(* IEC 61131-3 sources: NachHouse_TST/API/api_V12 (part 2) *)

(* ---- _07_RxBuf.ST ---- *)
// Limity jedného prijímacieho bloku a celého súboru ; Limits for one receive block and the complete file.
VAR_GLOBAL CONSTANT
  RB_BYTES {HIDDEN}    : UINT := 256;     // Maximálny počet dátových bajtov v jednom bloku ; Maximum data bytes in one block.
  RB_FILE_MAX {HIDDEN} : UDINT := 65535;  // Maximálna veľkosť súboru, ktorý možno zložiť ; Maximum size of a file that can be assembled.
END_VAR

VAR_GLOBAL
  RbSeen     : UDINT := 0;            // Posledná požiadavka bloku už prijatá PLC ; Most recent block request already consumed by the PLC.
  RbActive   : BOOL := FALSE;         // TRUE počas skladania viacerých blokov jedného súboru ; TRUE while assembling a file from multiple blocks.
  RbTotalW   : UDINT := 0;            // Očakávaná celková dĺžka aktuálneho súboru ; Expected total length of the current file.
  RbCrcW     : DWORD := 0;            // Očakávaný CRC32 súčet aktuálneho súboru ; Expected CRC32 checksum for the current file.
  RbCrcState : DWORD := 16#FFFFFFFF;  // Medzistav výpočtu CRC32 medzi prijatými blokmi ; Running CRC32 state across received blocks.
END_VAR

// Jeden krok štandardného CRC32 pre jeden bajt ; polynóm je 0xEDB88320. ; One standard CRC32 step for a byte ; the polynomial is 0xEDB88320.
// Pridá jeden bajt do priebežného výpočtu CRC32 ; Add one byte to the running CRC32 calculation.
FUNCTION RbCrcByte : DWORD
  VAR_INPUT
    State : DWORD;  // Doterajší priebežný stav CRC ; Previous running CRC state.
    B     : BYTE;   // Bajt, ktorý sa pridáva do CRC ; Byte to add to the CRC.
  END_VAR
  VAR
    C : DWORD;  // Pracovný 32-bitový stav CRC ; Working 32-bit CRC value.
    I : USINT;  // Počet ôsmich bitových krokov jedného bajtu ; Counter for the eight bit steps of one byte.
  END_VAR
  C := State XOR BYTE_TO_DWORD(B);
  FOR I := 1 TO 8 DO
    IF (C AND 16#00000001) <> 0 THEN
      C := SHR(C, 1) XOR 16#EDB88320;
    ELSE
      C := SHR(C, 1);
    END_IF;
  END_FOR;
  RbCrcByte := C;
END_FUNCTION

// Každé nové RbRq spracuje jeden blok ; RbAck potvrdí spracovanie a RbErr výsledok. ; Each new RbRq processes one block ; RbAck acknowledges it and RbErr reports the result.
// RbReady sa nastaví až po kontrole veľkosti a CRC celého súboru. ; RbReady is set only after validating the full file size and CRC.
// Pri novej RbRq zapíše jeden blok do rx.json, priebežne počíta CRC a potvrdí výsledok ; On a new RbRq, write one block to rx.json, update CRC, and acknowledge the result.
FUNCTION RbCycle : BOOL
  VAR
    Hnd      : HANDLE;       // Otvorený súborový handle pre zápis bloku ; File handle used to write the block.
    Mode     : TF_MODE;      // Režim otvorenia: nový súbor alebo pripojenie ďalšieho bloku ; Open mode: create a file or append the next block.
    N        : UDINT;        // Počet bajtov, ktoré FileWrite skutočne zapísal ; Number of bytes actually written by FileWrite.
    I        : UINT;         // Index bajtu pri aktualizácii CRC ; Byte index while updating the CRC.
    PB       : PTR_TO BYTE;  // Ukazovateľ na postupné čítanie bajtov z rxBuf ; Pointer used to read bytes sequentially from rxBuf.
    Closed   : BOOL;         // Výsledok uzatvorenia súboru po zápise ; Result of closing the file after writing.
    FinalCrc : DWORD;        // Dokončený CRC32 súčet po spracovaní posledného bajtu ; Final CRC32 value after the last byte.
  END_VAR
  RbCycle := TRUE;
  // Bez nového čísla požiadavky sa blok nespracúva znova ; Do not process a block again without a new request number.
  IF (RbRq = 0) OR (RbRq = RbSeen) THEN RETURN; END_IF;
  RbSeen := RbRq;
  RbErr := 0;

  // Počas parsovania JSON-u sa ďalší blok odmietne, aby sa súbor nemenil pod parserom ; Reject a new block while JSON parsing is active so the file cannot change underneath the parser.
  IF RxSt <> 0 THEN RbErr := 10;
  ELSIF (RbLen = 0) OR (RbLen > RB_BYTES) THEN RbErr := 1;
  ELSIF (RbTotal = 0) OR (RbTotal > RB_FILE_MAX) THEN RbErr := 2;
  ELSIF RbOfs > RbTotal THEN RbErr := 3;
  ELSIF UINT_TO_UDINT(RbLen) > RbTotal - RbOfs THEN RbErr := 3;
  END_IF;

  // Pokračuje iba po úspešných kontrolách dĺžky a rozsahu ; Continue only after length and range validation succeeds.
  IF RbErr = 0 THEN
    IF RbOfs = 0 THEN
      RbActive := TRUE;
      RbReady := FALSE;
      RbWrote := 0;
      RbTotalW := RbTotal;
      RbCrcW := RbCrc;
      RbCrcState := 16#FFFFFFFF;
      Mode := F_WRITE;
    ELSE
      Mode := F_APPEND;
      IF NOT RbActive THEN RbErr := 4;
      ELSIF RbOfs <> RbWrote THEN RbErr := 5;
      ELSIF (RbTotal <> RbTotalW) OR (RbCrc <> RbCrcW) THEN RbErr := 6;
      END_IF;
    END_IF;
  END_IF;

  // Pokračuje iba po úspešných kontrolách dĺžky a rozsahu ; Continue only after length and range validation succeeds.
  IF RbErr = 0 THEN
    Hnd := FileOpen(fileName := RxPath, mode := Mode);  // Otvorí rx.json na prvý zápis alebo doplnenie bloku ; Open rx.json for the first write or for appending a block.
    IF Hnd = INVALID_HANDLE_VALUE THEN
      RbErr := 7;
      RbActive := FALSE;
    ELSE
      N := FileWrite(hFile := Hnd, adrBuf := PTR_TO_UDINT(ADR(rxBuf[0])),
                     size := UINT_TO_UDINT(RbLen));
      Closed := FileClose(hFile := Hnd);
      IF (N <> UINT_TO_UDINT(RbLen)) OR NOT Closed THEN
        RbErr := 8;
        RbActive := FALSE;
      ELSE
        PB := ADR(rxBuf[0]);  // Začne kontrolný súčet od prvého bajtu aktuálneho bloku ; Start checksum calculation at the first byte of this block.
        FOR I := 1 TO RbLen DO
          RbCrcState := RbCrcByte(State := RbCrcState, B := PB^);
          PB := UDINT_TO_PTR(PTR_TO_UDINT(PB) + 1);
        END_FOR;
        RbWrote := RbWrote + UINT_TO_UDINT(RbLen);
        // Po prijatí deklarovaného počtu bajtov overí CRC celého súboru ; Once the declared byte count arrives, verify the complete-file CRC.
        IF RbWrote = RbTotalW THEN
          FinalCrc := RbCrcState XOR 16#FFFFFFFF;
          IF FinalCrc = RbCrcW THEN
            RbReady := TRUE;
          ELSE
            RbErr := 9;
          END_IF;
          RbActive := FALSE;
        END_IF;
      END_IF;
    END_IF;
  END_IF;

  RbAck := RbRq;  // Potvrdí spracovanie aj prípadnú chybu tohto bloku ; Acknowledge processing, including any block error.
  RbCycle := RbErr = 0;
END_FUNCTION

(* ---- _02_DataInit.ST ---- *)
// Naplní testovacie záznamy a jednorazovo ich skopíruje do mRam. ; Populate test records and copy them into mRam once.
// Pri prvom cykle vytvorí testovacie ROOM/USER dáta a skopíruje ich do mRam ; On the first cycle, creates test ROOM/USER data and copies it into mRam.
FUNCTION InitData : BOOL
  VAR
    Rec    : INT;    // Index testovanej vety 1..10 ; Test record index, 1..10.
    Pos    : INT;    // Index prvku vnútorného poľa používateľa ; Index into a nested user array.
    Copied : UDINT;  // Počet bajtov skutočne skopírovaných funkciou MemCpyPtr ; Number of bytes actually copied by MemCpyPtr.
  END_VAR
  InitData := TRUE;
  // Inicializáciu vykoná iba pri štartovacej hodnote Ini ; Initialize only when Ini has its startup value.
  IF aSys.Ini <> 250 THEN RETURN; END_IF;

  // Naplnenie desiatich testovacích viet oboch typov ; Fill ten test records for both data types.
  FOR Rec := 1 TO 10 DO
    yRooms[Rec].mem.rec.Ok := TRUE;  // Začiatok naplnenia stavovej a konfiguračnej časti aktuálnej miestnosti ; Begin filling the current room's state and configuration.
    yRooms[Rec].mem.rec.ID := Rec;
    yRooms[Rec].mem.all.RoomID := Rec;
    yRooms[Rec].mem.all.CategoryID := 5;
    yRooms[Rec].mem.Temperature := 20.0 + INT_TO_REAL(Rec);
    yRooms[Rec].mem.Humidity := 40.0 + INT_TO_REAL(Rec);
    yRooms[Rec].mem.Presence := (Rec MOD 2) = 0;
    yRooms[Rec].mem.DayPhase := INT_TO_UINT(140 + Rec);
    yRooms[Rec].mem.CategoryMask := 16#00000005;
    yRooms[Rec].mem.AlarmLevel := INT_TO_USINT(Rec MOD 3);
    yRooms[Rec].mem.Online := TRUE;
    yRooms[Rec].mem.Twilight := (Rec MOD 2) <> 0;
    yRooms[Rec].cfg.Name := 'Test room';
    yRooms[Rec].cfg._Dint := INT_TO_DINT(-1000 - Rec);
    yRooms[Rec].cfg._Sint := INT_TO_SINT(-10 + Rec);
    yRooms[Rec].cfg._Usint := INT_TO_USINT(100 + Rec);
    yRooms[Rec].cfg._Uint := INT_TO_UINT(1000 + Rec);
    yRooms[Rec].cfg._Real := 10.5 + INT_TO_REAL(Rec);
    yRooms[Rec].cfg._LReal := 1000.5 + INT_TO_LREAL(Rec);
    yRooms[Rec].cfg._String := '';
    yRooms[Rec].cfg._StringCZSK := 'SVKBEGIN_+ľščťžýáíé_SVKEND';
    yRooms[Rec].cfg._BYTE := 16#A5; yRooms[Rec].cfg._WORD := 16#A55A;
    yRooms[Rec].cfg._TIME := T#12h34m56s789ms;
    yRooms[Rec].cfg._DATE := D#2026-10-07;
    yRooms[Rec].cfg._TIME_OF_DAY := TOD#12:34:56.789;
    yRooms[Rec].cfg._DATE_AND_TIME := DT#2026-10-07-12:34:56.789;

    yUsers[Rec].mem.rec.Ok := TRUE; yUsers[Rec].mem.rec.ID := Rec;  // Začiatok naplnenia aktuálnej testovacej vety USER ; Begin filling the current USER test record.
    yUsers[Rec].mem.all.RoomID := Rec; yUsers[Rec].mem.all.CategoryID := 1;
    yUsers[Rec].mem.Connected := (Rec MOD 2) = 0;
    yUsers[Rec].mem.LastError := '';
    yUsers[Rec].mem.LastUpdate := UDINT#2026100700 + INT_TO_UDINT(Rec);
    yUsers[Rec].cfg.Name := 'Test user'; yUsers[Rec].cfg.LoginHome := TRUE;
    yUsers[Rec].cfg.DshSet := FALSE; yUsers[Rec].cfg.OwnDSH := TRUE;
    yUsers[Rec].cfg.OwnQCK := TRUE;
    yUsers[Rec].cfg.UsrRight := INT_TO_USINT(1 + (Rec MOD 3));
    // Zónové oprávnenia sa menia podľa čísla testovacej vety ; Zone permissions vary with the test-record number.
    FOR Pos := 1 TO 16 DO yUsers[Rec].cfg.ZonList[Pos] := Pos <= (Rec + 1); END_FOR;
    yUsers[Rec].cfg.sbj := INT_TO_USINT(Rec);
    yUsers[Rec].cfg.lng := INT_TO_USINT(Rec MOD 2);
    FOR Pos := 0 TO 7 DO
      yUsers[Rec].cfg.fav[Pos] := INT_TO_USINT(Pos + Rec);
      yUsers[Rec].cfg.msg[Pos] := Pos = (Rec MOD 8);
    END_FOR;
    yUsers[Rec].cfg.keyPas := '123456'; yUsers[Rec].cfg.IPnbr := 1;
    yUsers[Rec].cfg.IP[1] := '192.168.33.10';
    yUsers[Rec].cfg.IP[2] := ''; yUsers[Rec].cfg.IP[3] := '';
    yUsers[Rec].cfg.mail := 'test@example.com';
    yUsers[Rec].cfg.TOKENAPPLE := 'apple-test-token';
    yUsers[Rec].cfg.TOKENUNI := 'uni-test-token';
    yUsers[Rec].cfg.gsm := '+421900000000';
    yUsers[Rec].cfg.skin := INT_TO_USINT(Rec MOD 2);
    FOR Pos := 0 TO 30 DO
      IF Pos = 0 THEN yUsers[Rec].cfg.Brw[Pos] := 0;
      ELSE yUsers[Rec].cfg.Brw[Pos] := 1;
      END_IF;
    END_FOR;
  END_FOR;

  aCfg[1].iRam := 0;  // ROOM zaberá prvú oblasť mRam od bajtu nula ; ROOM occupies the first mRam region starting at byte zero.
  aCfg[2].iRam := aCfg[1].Siz * aCfg[1].Rec;  // USER oblasť začína bezprostredne za všetkými vetami ROOM ; USER starts immediately after all ROOM records.
  xRoom := ADR(mRam[aCfg[1].iRam]);  // Vypočíta ukazovateľ na prvú ROOM vetu ; Calculate a pointer to the first ROOM record.
  xUser := ADR(mRam[aCfg[2].iRam]);  // Vypočíta ukazovateľ na prvú USER vetu ; Calculate a pointer to the first USER record.
  aCfg[1].Ram := PTR_TO_UDINT(xRoom);  // Uloží absolútnu adresu ROOM oblasti pre adresovanie schémou ; Store the ROOM base address for schema-based access.
  aCfg[2].Ram := PTR_TO_UDINT(xUser);  // Uloží absolútnu adresu USER oblasti pre adresovanie schémou ; Store the USER base address for schema-based access.
  Copied := MemCpyPtr(source := ADR(yRooms[1]), dest := xRoom, length := aCfg[1].Siz * aCfg[1].Rec);  // Skopíruje všetkých desať testovacích miestností do súvislej oblasti mRam ; Copy all ten test rooms into their contiguous mRam region.
  aCfg[1].ok := Copied = aCfg[1].Siz * aCfg[1].Rec;
  Copied := MemCpyPtr(source := ADR(yUsers[1]), dest := xUser, length := aCfg[2].Siz * aCfg[2].Rec);  // Skopíruje všetkých desať testovacích používateľov do mRam ; Copy all ten test users into mRam.
  aCfg[2].ok := Copied = aCfg[2].Siz * aCfg[2].Rec;
  aSys.Restart := FALSE;  // Označí dokončenie štartovacej inicializácie ; Mark startup initialization as complete.
  aSys.Ini := 0;  // Zabráni opätovnému naplneniu testovacích dát v ďalších cykloch ; Prevent test data from being initialized again in later cycles.
END_FUNCTION

(* ---- prgMain.ST ---- *)
// Hlavný cyklický program: inicializácia, schéma, export, blokový príjem a import ; Main cyclic program: initialization, schema, export, block receive, and import.
PROGRAM prgMain
  VAR
    DepStarted  : BOOL := FALSE;  // Určuje, či sa vykonal úvodný reset požiadavky na balík ; Tracks whether the initial package-request reset has run.
    DepAccepted : BOOL;           // Pracovný výsledok prijatia balíka PLC ; Temporary result of PLC package acceptance.
  END_VAR

  InitData();  // Musí byť prvé: testovacie dáta a mRam sa inicializujú pred ostatnými cyklami. ; Keep this first: test data and mRam must be initialized before the other cycles.
  SchInit();  // Overí tabuľku schémy oproti typom a rozloženiu pamäte ; Validate the schema table against types and memory layout.
  TxCycle();  // Obslúži prípadnú požiadavku klienta na export JSON ; Process a client request to export JSON.
  RbCycle();  // Spracuje nový prijatý blok a prípadne doplní rx.json ; Process a new received block and append it to rx.json.
  RxCycle();  // Spracuje požiadavku na prevod rx.json do mRam ; Process a request to convert rx.json into mRam.

  IF NOT DepStarted THEN
    DepRq := FALSE;  // Počiatočne zruší požiadavku, aby sa nespustil nechcený deploy ; Clear the request initially to avoid an unintended deployment.
    DepRes := 0;
    DepStarted := TRUE;
  ELSIF DepRq THEN
    DepRq := FALSE;  // Zruší prijatú požiadavku pred načítaním balíka ; Clear the accepted request before loading the package.
    DepAccepted := LoadNewPackage2(rq := TRUE, pckg := '//WWW/UPLOAD/NEW_PACK.TTR');  // Požiada PLC o načítanie balíka z určeného súboru ; Ask the PLC to load the package from the specified file.
    // Vráti stav úspešného prijatia balíka ; Return the package-accepted status.
    IF DepAccepted THEN DepRes := 1;
    ELSE DepRes := 3;
    END_IF;
  END_IF;
END_PROGRAM
